(* IEC 61131-3 sources: SemantiST/compiler/toolchain/compatibility/profiles/codesys-memory, 1 file *)

(* ---- interfaces.st ---- *)
(* Deterministic CODESYS memory compatibility backed by runtime.c. *)

@EXTERNAL FUNCTION __SEMANTIST_MEMSET : REF_TO BYTE
VAR_INPUT
    DEST : REF_TO BYTE;
    VALUE : UDINT;
    COUNT : UDINT;
END_VAR
END_FUNCTION

@EXTERNAL FUNCTION __SEMANTIST_MEMCPY : REF_TO BYTE
VAR_INPUT
    DEST : REF_TO BYTE;
    SOURCE : REF_TO BYTE;
    COUNT : UDINT;
END_VAR
END_FUNCTION

@EXTERNAL FUNCTION __SEMANTIST_MEMMOVE : REF_TO BYTE
VAR_INPUT
    DEST : REF_TO BYTE;
    SOURCE : REF_TO BYTE;
    COUNT : UDINT;
END_VAR
END_FUNCTION

FUNCTION SysMemSet : REF_TO BYTE
VAR_INPUT
    pDest : REF_TO BYTE;
    udiValue : UDINT;
    udiCount : UDINT;
END_VAR
SysMemSet := __SEMANTIST_MEMSET(pDest, udiValue, udiCount);
END_FUNCTION

FUNCTION SysMemCpy : REF_TO BYTE
VAR_INPUT
    pDest : REF_TO BYTE;
    pSrc : REF_TO BYTE;
    udiCount : UDINT;
END_VAR
SysMemCpy := __SEMANTIST_MEMCPY(pDest, pSrc, udiCount);
END_FUNCTION

FUNCTION SysMemMove : REF_TO BYTE
VAR_INPUT
    pDest : REF_TO BYTE;
    pSrc : REF_TO BYTE;
    udiCount : UDINT;
END_VAR
SysMemMove := __SEMANTIST_MEMMOVE(pDest, pSrc, udiCount);
END_FUNCTION
